(* IEC 61131-3 sources: llm-plc-st-eval/data/definitivo/gemini-3.1-pro-preview/B3/few_shot, 3 files *)

(* ---- ejec_1.st ---- *)
FUNCTION_BLOCK FB_Contador
VAR_INPUT
    sensorPieza : BOOL; (* Sensor de deteccion de pieza *)
    btnReset : BOOL; (* Boton de reinicio *)
END_VAR
VAR_OUTPUT
    loteListo : BOOL; (* Salida de lote completo *)
    cuenta : INT; (* Cantidad de piezas contadas *)
END_VAR
VAR
    ctPiezas : CTU; (* Bloque contador ascendente *)
END_VAR

(* El contador incrementa con el flanco de subida del sensor *)
ctPiezas(CU := sensorPieza, R := btnReset, PV := 12);

(* Asignacion de salidas *)
loteListo := ctPiezas.Q;
cuenta := ctPiezas.CV;
END_FUNCTION_BLOCK

(* ---- ejec_2.st ---- *)
FUNCTION_BLOCK FB_Contador
VAR_INPUT
    sensorPieza : BOOL; (* Sensor fotoelectrico de piezas *)
    btnReset : BOOL; (* Boton de reinicio de cuenta *)
END_VAR
VAR_OUTPUT
    loteListo : BOOL; (* Indicador de lote completo *)
    cuenta : INT; (* Cantidad actual de piezas *)
END_VAR
VAR
    contador : CTU; (* Bloque contador ascendente *)
END_VAR

(* El contador incrementa con el flanco de subida del sensor y se reinicia con el boton *)
contador(CU := sensorPieza, RESET := btnReset, PV := 12);

(* Asignacion de salidas *)
loteListo := contador.Q;
cuenta := contador.CV;
END_FUNCTION_BLOCK

(* ---- ejec_3.st ---- *)
FUNCTION_BLOCK FB_Contador
VAR_INPUT
    sensorPieza : BOOL; (* Sensor de pieza *)
    btnReset : BOOL; (* Boton de reset *)
END_VAR
VAR_OUTPUT
    loteListo : BOOL; (* Salida de lote completo *)
    cuenta : INT; (* Cuenta de piezas *)
END_VAR
VAR
    cPiezas : CTU; (* Contador ascendente *)
END_VAR

(* Incrementa con cada pieza, activa salida al llegar a 12 y permite reset *)
cPiezas(CU := sensorPieza, RESET := btnReset, PV := 12);
loteListo := cPiezas.Q;
cuenta := cPiezas.CV;
END_FUNCTION_BLOCK
